Fanuc KAREL source: KT00975.KL

PROGRAM KT00975
%NOLOCKGROUP
VAR
  ENTRY: INTEGER
  PNAME: STRING[80]
  VNAME: STRING[80]
  STATUS: INTEGER
  VALUE: ARRAY[4] OF XYZWPR
BEGIN
  ENTRY = 0
  PNAME = ''
  VNAME = 'VALUE'
  SET_VAR(ENTRY, PNAME, VNAME, VALUE, STATUS)
END KT00975
